Fanuc KAREL source: kb00188.KL

-- PROVISIONAL review KL for V1013-1; original PC SHA256 6af46d9a7b4b1bc8b0618537e0fe70996a83ca9e8c419cf60959fd604fac3b3e
-- Incomplete behavior may be omitted. Consult companion uncertainty JSON. Do not deploy.
PROGRAM KB00188
%NOLOCKGROUP
VAR
  P1 : STRING[80]
  RESULT : INTEGER
BEGIN
  -- UNRESOLVED_PC offsets 5-14; opcodes 3F,75
  -- UNRESOLVED_PC offsets 19-36; opcodes 27,22,2A,76,23
  -- UNRESOLVED_PC offsets 41-45; opcodes 7F
END KB00188
